Fanuc KAREL source: kb00186.KL

-- PROVISIONAL review KL for V1013-1; original PC SHA256 6c2149964cff5216c5f6ee726e06d123303d80d20ac1bff2c56024dddd2d4ac7
-- Incomplete behavior may be omitted. Consult companion uncertainty JSON. Do not deploy.
PROGRAM KB00186
%NOLOCKGROUP
VAR
  P1 : REAL
  RESULT : REAL
BEGIN
  -- UNRESOLVED_PC offsets 5-16; opcodes 2E,23
  -- UNRESOLVED_PC offsets 21-36; opcodes 27,22,76,23
  -- UNRESOLVED_PC offsets 41-45; opcodes 7F
END KB00186
